TYPE ST_EL3312CoeInfo :
STRUCT
	bEnableUserScale 			:BOOL := FALSE;
	bEnableFilter 					:BOOL := FALSE;
	bEnableLimit1 				:BOOL := FALSE;
	bEnableLimit2 				:BOOL := FALSE;
	bEnableUserCalibration 		:BOOL := FALSE;
	bEnableVendorCalibration 		:BOOL := TRUE;
	dwColdjunctionCompensation 	:DWORD := 0;
	nUserScaleOffset 				:INT := 0;
	dnUserScaleGain 				:DINT := 65536;
	nLimit1 						:INT := 0;
	nLimit2 						:INT := 0;
	dwFilterSettings 				:DWORD := 0;
	nUserCalibrationOffset 			:INT := 0;
	unUserCalibrationGain 			:UINT := 65535;
	dwTCElement 				:DWORD := 0;
END_STRUCT
END_TYPE

(* stored: Version 1.1.0.1, ProductVersion 3.1.4024.15
   DUT ST_EL3312CoeInfo: Id {adee76d3-de0d-4329-ae4b-889034468403} *)
